FUNCTION_BLOCK IOTest16 (* CAT Function Block Type *)
  (* Standard: 61499-2 *)
  (* Version 0.0, 11/13/2026, Sandeep Patil, Flexbridge AB, template *)
  PACKAGE Flexbridge.FestoMPS400;
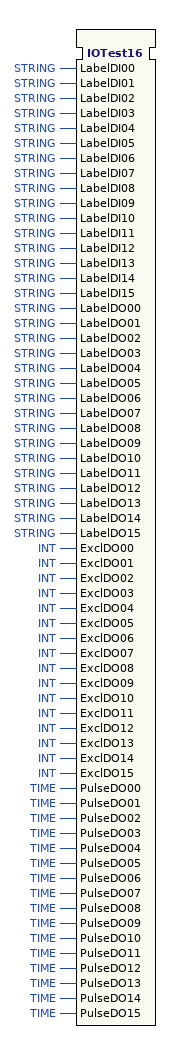
  VAR_INPUT
    LabelDI00 : STRING; (* Text next to input lamp 00 *)
    LabelDI01 : STRING; (* Text next to input lamp 01 *)
    LabelDI02 : STRING; (* Text next to input lamp 02 *)
    LabelDI03 : STRING; (* Text next to input lamp 03 *)
    LabelDI04 : STRING; (* Text next to input lamp 04 *)
    LabelDI05 : STRING; (* Text next to input lamp 05 *)
    LabelDI06 : STRING; (* Text next to input lamp 06 *)
    LabelDI07 : STRING; (* Text next to input lamp 07 *)
    LabelDI08 : STRING; (* Text next to input lamp 08 *)
    LabelDI09 : STRING; (* Text next to input lamp 09 *)
    LabelDI10 : STRING; (* Text next to input lamp 10 *)
    LabelDI11 : STRING; (* Text next to input lamp 11 *)
    LabelDI12 : STRING; (* Text next to input lamp 12 *)
    LabelDI13 : STRING; (* Text next to input lamp 13 *)
    LabelDI14 : STRING; (* Text next to input lamp 14 *)
    LabelDI15 : STRING; (* Text next to input lamp 15 *)
    LabelDO00 : STRING; (* Text on output button 00 *)
    LabelDO01 : STRING; (* Text on output button 01 *)
    LabelDO02 : STRING; (* Text on output button 02 *)
    LabelDO03 : STRING; (* Text on output button 03 *)
    LabelDO04 : STRING; (* Text on output button 04 *)
    LabelDO05 : STRING; (* Text on output button 05 *)
    LabelDO06 : STRING; (* Text on output button 06 *)
    LabelDO07 : STRING; (* Text on output button 07 *)
    LabelDO08 : STRING; (* Text on output button 08 *)
    LabelDO09 : STRING; (* Text on output button 09 *)
    LabelDO10 : STRING; (* Text on output button 10 *)
    LabelDO11 : STRING; (* Text on output button 11 *)
    LabelDO12 : STRING; (* Text on output button 12 *)
    LabelDO13 : STRING; (* Text on output button 13 *)
    LabelDO14 : STRING; (* Text on output button 14 *)
    LabelDO15 : STRING; (* Text on output button 15 *)
    ExclDO00 : INT := -1; (* Output that must never be on together with output 00; -1 = none *)
    ExclDO01 : INT := -1; (* Output that must never be on together with output 01; -1 = none *)
    ExclDO02 : INT := -1; (* Output that must never be on together with output 02; -1 = none *)
    ExclDO03 : INT := -1; (* Output that must never be on together with output 03; -1 = none *)
    ExclDO04 : INT := -1; (* Output that must never be on together with output 04; -1 = none *)
    ExclDO05 : INT := -1; (* Output that must never be on together with output 05; -1 = none *)
    ExclDO06 : INT := -1; (* Output that must never be on together with output 06; -1 = none *)
    ExclDO07 : INT := -1; (* Output that must never be on together with output 07; -1 = none *)
    ExclDO08 : INT := -1; (* Output that must never be on together with output 08; -1 = none *)
    ExclDO09 : INT := -1; (* Output that must never be on together with output 09; -1 = none *)
    ExclDO10 : INT := -1; (* Output that must never be on together with output 10; -1 = none *)
    ExclDO11 : INT := -1; (* Output that must never be on together with output 11; -1 = none *)
    ExclDO12 : INT := -1; (* Output that must never be on together with output 12; -1 = none *)
    ExclDO13 : INT := -1; (* Output that must never be on together with output 13; -1 = none *)
    ExclDO14 : INT := -1; (* Output that must never be on together with output 14; -1 = none *)
    ExclDO15 : INT := -1; (* Output that must never be on together with output 15; -1 = none *)
    PulseDO00 : TIME := T#0s; (* Pulse time of output 00; T#0s = toggle *)
    PulseDO01 : TIME := T#0s; (* Pulse time of output 01; T#0s = toggle *)
    PulseDO02 : TIME := T#0s; (* Pulse time of output 02; T#0s = toggle *)
    PulseDO03 : TIME := T#0s; (* Pulse time of output 03; T#0s = toggle *)
    PulseDO04 : TIME := T#0s; (* Pulse time of output 04; T#0s = toggle *)
    PulseDO05 : TIME := T#0s; (* Pulse time of output 05; T#0s = toggle *)
    PulseDO06 : TIME := T#0s; (* Pulse time of output 06; T#0s = toggle *)
    PulseDO07 : TIME := T#0s; (* Pulse time of output 07; T#0s = toggle *)
    PulseDO08 : TIME := T#0s; (* Pulse time of output 08; T#0s = toggle *)
    PulseDO09 : TIME := T#0s; (* Pulse time of output 09; T#0s = toggle *)
    PulseDO10 : TIME := T#0s; (* Pulse time of output 10; T#0s = toggle *)
    PulseDO11 : TIME := T#0s; (* Pulse time of output 11; T#0s = toggle *)
    PulseDO12 : TIME := T#0s; (* Pulse time of output 12; T#0s = toggle *)
    PulseDO13 : TIME := T#0s; (* Pulse time of output 13; T#0s = toggle *)
    PulseDO14 : TIME := T#0s; (* Pulse time of output 14; T#0s = toggle *)
    PulseDO15 : TIME := T#0s; (* Pulse time of output 15; T#0s = toggle *)
  END_VAR
  (* 0 - INITIALIZATION *)
  (* 6 - HMI INTERFACE *)
  (* 1 - FUNCTIONAL INPUT INTERFACE (labels, exclusive pairs, pulse times) *)
  (* 5 - LOGICS *)
  (* 3 - FIELD INTERFACE (DI00-DI15 from the input module, DO00-DO15 to the output module) *)
  FBS
    EVENTCHAIN : EVENTCHAIN(NAME := 'APP_INIT', PRIO := 20);
    IThis : IOTest16_HMI(QI := TRUE);
    Logic : IOTest16Logic;
    PulseTimer : E_DELAY;
    DI00 : dISignal(Name := '$${PATH}DIn');
    DO00 : dOSignal(Name := '$${PATH}DOut');
    DI01 : dISignal(Name := '$${PATH}DIn');
    DO01 : dOSignal(Name := '$${PATH}DOut');
    DI02 : dISignal(Name := '$${PATH}DIn');
    DO02 : dOSignal(Name := '$${PATH}DOut');
    DI03 : dISignal(Name := '$${PATH}DIn');
    DO03 : dOSignal(Name := '$${PATH}DOut');
    DI04 : dISignal(Name := '$${PATH}DIn');
    DO04 : dOSignal(Name := '$${PATH}DOut');
    DI05 : dISignal(Name := '$${PATH}DIn');
    DO05 : dOSignal(Name := '$${PATH}DOut');
    DI06 : dISignal(Name := '$${PATH}DIn');
    DO06 : dOSignal(Name := '$${PATH}DOut');
    DI07 : dISignal(Name := '$${PATH}DIn');
    DO07 : dOSignal(Name := '$${PATH}DOut');
    DI08 : dISignal(Name := '$${PATH}DIn');
    DO08 : dOSignal(Name := '$${PATH}DOut');
    DI09 : dISignal(Name := '$${PATH}DIn');
    DO09 : dOSignal(Name := '$${PATH}DOut');
    DI10 : dISignal(Name := '$${PATH}DIn');
    DO10 : dOSignal(Name := '$${PATH}DOut');
    DI11 : dISignal(Name := '$${PATH}DIn');
    DO11 : dOSignal(Name := '$${PATH}DOut');
    DI12 : dISignal(Name := '$${PATH}DIn');
    DO12 : dOSignal(Name := '$${PATH}DOut');
    DI13 : dISignal(Name := '$${PATH}DIn');
    DO13 : dOSignal(Name := '$${PATH}DOut');
    DI14 : dISignal(Name := '$${PATH}DIn');
    DO14 : dOSignal(Name := '$${PATH}DOut');
    DI15 : dISignal(Name := '$${PATH}DIn');
    DO15 : dOSignal(Name := '$${PATH}DOut');
  END_FBS
  EVENT_CONNECTIONS
    EVENTCHAIN.EO TO IThis.B63507A5491DBA4C;
    IThis.64A629998C2B4D18 TO Logic.C8E24F7DFBF9DC0B;
    Logic.43EC3925751B5FC3 TO IThis.76823A330AA1E11A;
    Logic.43EC3925751B5FC3 TO EVENTCHAIN.ACK;
    IThis.46C3A447E157753C TO Logic.4F41D35F800CFC8F;
    IThis.28B4B8110E8B23BA TO Logic.A50B78E1728D04A4;
    Logic.95657124D8C8D43B TO IThis.54230140E274F0DB;
    Logic.34AB0D5D62F7B6BD TO IThis.34403BA68899974A;
    Logic.2259194325478FA9 TO PulseTimer.START;
    Logic.AF504EDCD2D79B37 TO PulseTimer.STOP;
    PulseTimer.EO TO Logic.3BECA61FDE7B44FF;
    DI00.CNF TO Logic.37D8E079D482C806;
    DI01.CNF TO Logic.37D8E079D482C806;
    DI02.CNF TO Logic.37D8E079D482C806;
    DI03.CNF TO Logic.37D8E079D482C806;
    DI04.CNF TO Logic.37D8E079D482C806;
    DI05.CNF TO Logic.37D8E079D482C806;
    DI06.CNF TO Logic.37D8E079D482C806;
    DI07.CNF TO Logic.37D8E079D482C806;
    DI08.CNF TO Logic.37D8E079D482C806;
    DI09.CNF TO Logic.37D8E079D482C806;
    DI10.CNF TO Logic.37D8E079D482C806;
    DI11.CNF TO Logic.37D8E079D482C806;
    DI12.CNF TO Logic.37D8E079D482C806;
    DI13.CNF TO Logic.37D8E079D482C806;
    DI14.CNF TO Logic.37D8E079D482C806;
    DI15.CNF TO Logic.37D8E079D482C806;
    Logic.51822766C426B5C0 TO DO00.REQ;
    Logic.51822766C426B5C0 TO DO01.REQ;
    Logic.51822766C426B5C0 TO DO02.REQ;
    Logic.51822766C426B5C0 TO DO03.REQ;
    Logic.51822766C426B5C0 TO DO04.REQ;
    Logic.51822766C426B5C0 TO DO05.REQ;
    Logic.51822766C426B5C0 TO DO06.REQ;
    Logic.51822766C426B5C0 TO DO07.REQ;
    Logic.51822766C426B5C0 TO DO08.REQ;
    Logic.51822766C426B5C0 TO DO09.REQ;
    Logic.51822766C426B5C0 TO DO10.REQ;
    Logic.51822766C426B5C0 TO DO11.REQ;
    Logic.51822766C426B5C0 TO DO12.REQ;
    Logic.51822766C426B5C0 TO DO13.REQ;
    Logic.51822766C426B5C0 TO DO14.REQ;
    Logic.51822766C426B5C0 TO DO15.REQ;
  END_CONNECTIONS
  DATA_CONNECTIONS
    LabelDI00 TO IThis.AAD360AE0031FBA7;
    LabelDI01 TO IThis.34F8F4E8D5BD5270;
    LabelDI02 TO IThis.711E2B78537B9C76;
    LabelDI03 TO IThis.EA5F92EF2702E72A;
    LabelDI04 TO IThis.B76F7352E26DAEE5;
    LabelDI05 TO IThis.0D90E8F0FD1572E3;
    LabelDI06 TO IThis.E6E724C318C07961;
    LabelDI07 TO IThis.FF560F6D08B1558D;
    LabelDI08 TO IThis.33F536C3388479B8;
    LabelDI09 TO IThis.0092EBF7D09B1BB1;
    LabelDI10 TO IThis.DFB9DE52D9D3F241;
    LabelDI11 TO IThis.F80C75F157269E73;
    LabelDI12 TO IThis.3A2AF3DB14E057B8;
    LabelDI13 TO IThis.696BAC93C6231267;
    LabelDI14 TO IThis.BE7DD780B388821F;
    LabelDI15 TO IThis.00B4737EF87E9111;
    LabelDO00 TO IThis.C91F03C5F3D96794;
    LabelDO01 TO IThis.6C3353A6278F31A7;
    LabelDO02 TO IThis.9A90B29082BAD88B;
    LabelDO03 TO IThis.DA1A96FCDFEEF866;
    LabelDO04 TO IThis.215A0125F98E8D42;
    LabelDO05 TO IThis.BE06B8F15663C0B1;
    LabelDO06 TO IThis.6305E534B39F2EE6;
    LabelDO07 TO IThis.89781FCD347D10FA;
    LabelDO08 TO IThis.84372BA8D08A8AC4;
    LabelDO09 TO IThis.D28F405939B8975E;
    LabelDO10 TO IThis.6B71D2D92FFB8089;
    LabelDO11 TO IThis.BF8ECB0CDB9E1E69;
    LabelDO12 TO IThis.6A2AD1AEF0A7089C;
    LabelDO13 TO IThis.3E5EF677AEEB17E9;
    LabelDO14 TO IThis.AD9EF1048BD1ACBA;
    LabelDO15 TO IThis.192C79BC3C368A07;
    ExclDO00 TO Logic.DDAE9F07F58D3AF3;
    ExclDO01 TO Logic.D490237C6D4E6516;
    ExclDO02 TO Logic.E50209420C009F4D;
    ExclDO03 TO Logic.A2672ABC3CF05A06;
    ExclDO04 TO Logic.A05A62EB81F65CCD;
    ExclDO05 TO Logic.B3814EB203391BC5;
    ExclDO06 TO Logic.99EC20DF40F4004D;
    ExclDO07 TO Logic.539F691D9B0278AE;
    ExclDO08 TO Logic.E5B6E21CFC3AC94B;
    ExclDO09 TO Logic.B9844DC9EC2DA2D3;
    ExclDO10 TO Logic.D8E968D9ED6EAD78;
    ExclDO11 TO Logic.BD42D8EE1CF28EC7;
    ExclDO12 TO Logic.8ABE4B38E6F4FDE1;
    ExclDO13 TO Logic.1B8E5A84135FAAE2;
    ExclDO14 TO Logic.59086C3BA1BC429D;
    ExclDO15 TO Logic.0A12E6B7B932122B;
    PulseDO00 TO Logic.E9B291DAE8EC3101;
    PulseDO01 TO Logic.7A512D95D4D0A61F;
    PulseDO02 TO Logic.7525532A8E06D4CE;
    PulseDO03 TO Logic.20EE2114B0F6DEE5;
    PulseDO04 TO Logic.715C126EE559FCC9;
    PulseDO05 TO Logic.F1A616C66D70ACBF;
    PulseDO06 TO Logic.D0FF2731166DFF80;
    PulseDO07 TO Logic.44692470B3E913D9;
    PulseDO08 TO Logic.7E55167A22BDC761;
    PulseDO09 TO Logic.B7057C48294FDC9E;
    PulseDO10 TO Logic.655342177DFDBEE1;
    PulseDO11 TO Logic.5E0272D074046E45;
    PulseDO12 TO Logic.99E7F0AA334970C5;
    PulseDO13 TO Logic.37A96D725CFAB133;
    PulseDO14 TO Logic.3223EB9B0F78537C;
    PulseDO15 TO Logic.03045199FBDEE93E;
    IThis.5894EF1F76DACBEF TO Logic.0EDDD3C97AD8F01D;
    IThis.0210C65D19A82559 TO Logic.B9E6EF29DE219689;
    IThis.680269FA2EA04FD1 TO Logic.B813F17B6064C18A;
    IThis.35D3947E2ABD81D4 TO Logic.1ECD9FF20E604D7E;
    IThis.4F8A76D29C6427F5 TO Logic.0889FE27E9AC83E5;
    IThis.34E981D743B5E114 TO Logic.9074CB2F470CFAB6;
    IThis.A4E053B122E4DEFE TO Logic.A3D544F56D200CE3;
    IThis.B46E07C375751ECD TO Logic.10748F208DCC929B;
    IThis.03FAD46C5D8D1BB6 TO Logic.8FBB0D2B7E3D4228;
    IThis.D33DD8C84FDCD9A9 TO Logic.3ACE7EDDDACA5682;
    IThis.AF4F70D66078F64D TO Logic.1351E0491AD76222;
    IThis.80C2EAF9C573BE9F TO Logic.A3712C3A94CC2AB6;
    IThis.BB4ED98C4E679B32 TO Logic.7829DE08B48CBA69;
    IThis.F53FDC552BC54BC6 TO Logic.9D95F0AA02B53062;
    IThis.28D6362AB72212B7 TO Logic.470106CE276F2006;
    IThis.30DBE17A2158E4C0 TO Logic.8D7AF47444EF7843;
    DI00.Out TO Logic.E88733B66EEDE5AC;
    DI01.Out TO Logic.2D9172D0E7F74B4A;
    DI02.Out TO Logic.2413D9E06A0A664C;
    DI03.Out TO Logic.229FEA2BAA13F955;
    DI04.Out TO Logic.8AE96DD03FA39359;
    DI05.Out TO Logic.9B9AF66C91608DD0;
    DI06.Out TO Logic.4B59957A10E9D2A8;
    DI07.Out TO Logic.92EC702D9FE9D6FB;
    DI08.Out TO Logic.1A3DAD59292D205F;
    DI09.Out TO Logic.6998087FAC67F3DD;
    DI10.Out TO Logic.753A90A42240AB8C;
    DI11.Out TO Logic.FDC421EAFC181624;
    DI12.Out TO Logic.0BE32C4A5AD3A5ED;
    DI13.Out TO Logic.E508BA5ACAC55AE7;
    DI14.Out TO Logic.C23C564628BECC7A;
    DI15.Out TO Logic.49E71BE0894ECE8C;
    Logic.04664C0CBB69D8D5 TO DO00.Signal;
    Logic.89A51AF88B7AA097 TO DO01.Signal;
    Logic.3AB76BADE1F2940E TO DO02.Signal;
    Logic.D70803A3D192B869 TO DO03.Signal;
    Logic.78B1306E37D3C554 TO DO04.Signal;
    Logic.A3E89E8867874630 TO DO05.Signal;
    Logic.334B40A2F4D71B13 TO DO06.Signal;
    Logic.DE950EAA1286FE39 TO DO07.Signal;
    Logic.CE47C34426EFB090 TO DO08.Signal;
    Logic.A413288515257406 TO DO09.Signal;
    Logic.C2357E05B78CD97A TO DO10.Signal;
    Logic.BE8E59BD43C3FE78 TO DO11.Signal;
    Logic.E286D5C4FA1ECD64 TO DO12.Signal;
    Logic.04A1CE1AF5BB5C0C TO DO13.Signal;
    Logic.D31B2FDCBDE9B579 TO DO14.Signal;
    Logic.A85E311937FF6E1C TO DO15.Signal;
    Logic.4B5EC8A5B332C6E6 TO IThis.D8822B67D02F9092;
    Logic.36A460996A9CEBAA TO IThis.5FCEC26253E236DD;
    Logic.EEEFA62CB9FCB4DC TO IThis.B6265428486F3C44;
    Logic.93D8556D9BF5BEDE TO IThis.350803B156590673;
    Logic.06DFEB3EA6402D6A TO IThis.08D042CA123BBAD6;
    Logic.847650F12A885802 TO IThis.CCBF62D8F886AF7C;
    Logic.AAC103CA2E5BE052 TO IThis.D19743C15D298BBE;
    Logic.447D9C7678504652 TO IThis.3E78C72AA8E3D7CE;
    Logic.E16DCAC5E8025B8F TO IThis.944F09A1740ED60C;
    Logic.B6CEDB756BE42D88 TO IThis.19911228B40C640C;
    Logic.8DB923E5026BA397 TO IThis.ADE63BA19C92226A;
    Logic.0EDCD0AE06406A09 TO IThis.A626A0A5B091DAA5;
    Logic.F94D2283B770D8ED TO IThis.04C923A6ED5ACDAD;
    Logic.DA0A6CF8ADAD5257 TO IThis.AABBB683BD394519;
    Logic.0AD975F74C991833 TO IThis.250639C9D2AC2F88;
    Logic.4815DE5BF679E0A9 TO IThis.521435408CEF7A3E;
    Logic.70542509E2B5733D TO IThis.E09A83D8A036E0B5;
    Logic.124542E49CA6AA23 TO IThis.AB87D38FEB7AD14B;
    Logic.0C4C190DABE52E6E TO IThis.CF1768B1C1E14D27;
    Logic.5FEB31C180EEE23E TO IThis.A2264B1337E3CE4F;
    Logic.B77A123416E9E838 TO IThis.5A3733277ADA1972;
    Logic.ABAB61C97C68E080 TO IThis.9ACC547135D942C2;
    Logic.3A934E9EBE304B9F TO IThis.F4751479B8EF136F;
    Logic.691E069AE5B99296 TO IThis.F3D21410B005D7DD;
    Logic.2EE13BAB9E6BB6F9 TO IThis.870CA74D6592AE8C;
    Logic.877766A2EA3666A1 TO IThis.76D1F83FA874663D;
    Logic.2909F54A051FC588 TO IThis.BBC6AFF2758488E3;
    Logic.0A8D17318C17F619 TO IThis.E6FB069BD7AE847F;
    Logic.F832BB0B12B6DF77 TO IThis.C65E5D253AE76FB6;
    Logic.BEF94186384B2688 TO IThis.4B9EB0BE8906812E;
    Logic.9475C4ECC76ECBAE TO IThis.5940D288A5435331;
    Logic.840AB1AF61ACDCBF TO IThis.1B42CA3924E970A2;
    Logic.6D052A3B40885921 TO IThis.E942C3278740B311;
    Logic.D2A00432A826B8DE TO IThis.2C7D3EFEDD65334C;
    Logic.074568EE3A022E5C TO IThis.218682D551B5E363;
    Logic.4A0020CA77DCD6AE TO IThis.BE9EA829314C321C;
    Logic.218A6BCF580FB933 TO IThis.1A6032D49A7418F6;
    Logic.5125227FF732F976 TO IThis.5CFB3642C430CA38;
    Logic.74FA905002DF3FC5 TO IThis.DFD7541C44C59897;
    Logic.49A280672D3D265F TO IThis.C3C6D2AF4F6B5A2B;
    Logic.B30658EF959D2757 TO IThis.46D1595BC77B5B44;
    Logic.3AA55A681C7F4560 TO IThis.6375DB34DE05CEDB;
    Logic.B5C9E4089E02069C TO IThis.223D8DD33D7A9374;
    Logic.FA55C4B1BDFCF1FF TO IThis.73CF9439ACCA3B49;
    Logic.6016850F89DCAD9B TO IThis.CC9913EA3EC62326;
    Logic.D1EE8ED0B0C69C1A TO IThis.F4C67A480DCCD141;
    Logic.C416F1247A07DDE9 TO IThis.9EC199434FC33EAC;
    Logic.D280A15AC902A5AE TO IThis.C2165E4B8F3E9590;
    Logic.FEFD9E0A876A54DD TO PulseTimer.DT;
  END_CONNECTIONS
END_FUNCTION_BLOCK
